Staubli VAL3: loadSAFE.pgx

public program loadSAFE(num x_nLib, num& x_nResult)
  local string l_sPath
begin
  l_sPath="Disk://data/CustomerLib/lib"+toString("",x_nLib)+"/safeData/safeData.pjx"
  x_nResult=safeTemp:libLoad(l_sPath)
  delay(0)
  logMsg(toString("",x_nResult))
end
